// TIA Portal V20 export
// export: Created 2026-10-19T18:45:50.3471132Z, ExportSetting None, DisplayName Totally Integrated Automation Portal, DisplayVersion V20 Update 6, DisplayName TIA Portal Openness, DisplayVersion V20 Update 6, DisplayName TIA Portal Version Control Interface, DisplayVersion V20 Update 6, DisplayName SINAMICS Startdrive Advanced, DisplayVersion V20 SP1, DisplayName SINAMICS Startdrive G130, G150, S120, S150, SINAMICS MV, G220, S200, S210, DisplayVersion V20 SP1, DisplayName SINAMICS Startdrive G110M, G120, G120C, G120D, G120P, G115D, DisplayVersion V20 SP1, DisplayName STEP 7 Professional, DisplayVersion V20 Update 6, DisplayName STEP 7 Safety, DisplayVersion V20 Update 2, DisplayName WinCC Basic/Comfort/Advanced, DisplayVersion V20 Update 6, DisplayName WinCC Unified, DisplayVersion V20 Update 6
VAR_GLOBAL   // PLC tag table "IO_Charger Panel_L4"
   "CHARGER L4 - Output Voltage" AT %ID828 : Real;   // Actual Output Voltage
   "CHARGER L4 - Output Current" AT %ID832 : Real;   // Actual Output Current
   "CHARGER L4 - Set Voltage Feedback" AT %ID836 : Real;   // Set Voltage Value
   "CHARGER L4 - Set Current Feedback" AT %ID840 : Real;   // Set Current Value
   "CHARGER L4 - Charging Start" AT %I848.0 : Bool;   // Charging Running Status
   "CHARGER L4 - Set Voltage Output" AT %QD414 : Real;   // Issue Target Voltage
   "CHARGER L4 - Set Current Output" AT %QD418 : Real;   // Issue Target Current
   "CHARGER L4 - Start Charging" AT %Q422.0 : Bool;   // Start Charging Command
   "CHARGER L4 - Stop Charging" AT %Q422.1 : Bool;   // Stop Charging Command
   "CHARGER L4 - Confirm Voltage & Current Setting" AT %Q422.2 : Bool;   // Confirmation Command
END_VAR
